(* IEC 61131-3 sources: llm-plc-st-eval/codesys/dobles/B4, 5 files *)

(* ---- 01_Correcta.st ---- *)
(* DOBLE DE PRUEBA B4/Correcta - NO ES CORPUS. Esperado: veredicto 1 *)
FUNCTION_BLOCK FB_Giro
VAR_INPUT
    btnFwd : BOOL;
    btnRev : BOOL;
    btnParo : BOOL;
END_VAR
VAR_OUTPUT
    fwd : BOOL;
    rev : BOOL;
END_VAR
VAR
    nada : BOOL;
END_VAR
IF btnParo THEN
    fwd := FALSE;
    rev := FALSE;
ELSE
    IF btnFwd AND NOT rev THEN
        fwd := TRUE;
    END_IF
    IF btnRev AND NOT fwd THEN
        rev := TRUE;
    END_IF
END_IF
END_FUNCTION_BLOCK

(* ---- 02_SinEnclavamiento.st ---- *)
(* DOBLE DE PRUEBA B4/SinEnclavamiento - NO ES CORPUS. Esperado: veredicto 2, falla en el paso 2 *)
FUNCTION_BLOCK FB_Giro
VAR_INPUT
    btnFwd : BOOL;
    btnRev : BOOL;
    btnParo : BOOL;
END_VAR
VAR_OUTPUT
    fwd : BOOL;
    rev : BOOL;
END_VAR
VAR
    nada : BOOL;
END_VAR
fwd := btnFwd AND NOT btnParo AND NOT btnRev;
rev := btnRev AND NOT btnParo AND NOT btnFwd;
END_FUNCTION_BLOCK

(* ---- 03_InversionDirecta.st ---- *)
(* DOBLE DE PRUEBA B4/InversionDirecta - NO ES CORPUS. Esperado: veredicto 2, falla en el paso 3 *)
FUNCTION_BLOCK FB_Giro
VAR_INPUT
    btnFwd : BOOL;
    btnRev : BOOL;
    btnParo : BOOL;
END_VAR
VAR_OUTPUT
    fwd : BOOL;
    rev : BOOL;
END_VAR
VAR
    nada : BOOL;
END_VAR
IF btnParo THEN
    fwd := FALSE;
    rev := FALSE;
ELSIF btnFwd THEN
    fwd := TRUE;
    rev := FALSE;
ELSIF btnRev THEN
    rev := TRUE;
    fwd := FALSE;
END_IF
END_FUNCTION_BLOCK

(* ---- 04_SinInterlock.st ---- *)
(* DOBLE DE PRUEBA B4/SinInterlock - NO ES CORPUS. Esperado: veredicto 2 *)
FUNCTION_BLOCK FB_Giro
VAR_INPUT
    btnFwd : BOOL;
    btnRev : BOOL;
    btnParo : BOOL;
END_VAR
VAR_OUTPUT
    fwd : BOOL;
    rev : BOOL;
END_VAR
VAR
    nada : BOOL;
END_VAR
IF btnParo THEN
    fwd := FALSE;
    rev := FALSE;
ELSE
    IF btnFwd THEN
        fwd := TRUE;
    END_IF
    IF btnRev THEN
        rev := TRUE;
    END_IF
END_IF
END_FUNCTION_BLOCK

(* ---- 05_CarreraDeInterlock.st ---- *)
(* DOBLE DE PRUEBA B4/CarreraDeInterlock - NO ES CORPUS. Esperado: veredicto 2 *)
FUNCTION_BLOCK FB_Giro
VAR_INPUT
    btnFwd : BOOL;
    btnRev : BOOL;
    btnParo : BOOL;
END_VAR
VAR_OUTPUT
    fwd : BOOL;
    rev : BOOL;
END_VAR
VAR
    fwdPrev : BOOL;
    revPrev : BOOL;
END_VAR
IF btnParo THEN
    fwd := FALSE;
    rev := FALSE;
ELSE
    IF btnFwd AND NOT revPrev THEN
        fwd := TRUE;
    END_IF
    IF btnRev AND NOT fwdPrev THEN
        rev := TRUE;
    END_IF
END_IF
fwdPrev := fwd;
revPrev := rev;
END_FUNCTION_BLOCK
